(* IEC 61131-3 sources: plcassist-cli/packages/volt-lsp-iec/test-corpus/lenze-mid/Device/Plc Logic/Application/Library Manager/CommFB, 41 files *)

(* ---- ADDRESSCONCEPT.gvl ---- *)
VAR_GLOBAL
	DUMMY : UDINT := 0;
END_VAR

(* ---- CONSTANTS.gvl ---- *)
VAR_GLOBAL
	INVALID_ID : UDINT := 16#FFFFFFFF;
	MAX_PN_ALARM_DATA : UDINT := 198;
END_VAR

(* ---- ICOMMFBALARMSENDER.itf ---- *)
INTERFACE ICOMMFBALARMSENDER
END_INTERFACE

METHOD ALARMCNF
VAR_INPUT
	ERROR : DWORD;
END_VAR
END_METHOD

(* ---- ICOMMFBCONNECTIONMANAGERFACTORY.itf ---- *)
INTERFACE ICOMMFBCONNECTIONMANAGERFACTORY
END_INTERFACE

METHOD GETCONNECTIONMANAGER : UDINT
VAR_INPUT
	CLIENT : IConnectionManagerClient;
END_VAR
VAR_OUTPUT
	CONNECTIONMANAGER : IConnectionManager;
END_VAR
VAR_IN_OUT
	D_ADDR : ADDR_TYPE;
END_VAR
END_METHOD

METHOD RELEASECONNECTIONMANAGER : UDINT
VAR_INPUT
	CLIENT : IConnectionManagerClient;
	CONNECTIONMANAGER : IConnectionManager;
END_VAR
END_METHOD

(* ---- ICOMMFBDIAGPROVIDER.itf ---- *)
INTERFACE ICOMMFBDIAGPROVIDER
END_INTERFACE

METHOD CHECKOWNER : BOOL
VAR_INPUT
	ID : UDINT;
END_VAR
END_METHOD

METHOD GETALARM : DWORD
VAR_INPUT
	MODE : INT;
	F_ID : DWORD;
END_VAR
VAR_OUTPUT
	NEW : BOOL;
	ID : DWORD;
	LEN : INT;
END_VAR
VAR_IN_OUT
	AINFO : AINFO_TYPE;
	CURRENTALARMID : UDINT;
END_VAR
END_METHOD

METHOD GETDIAG : DWORD
VAR_INPUT
	ID : DWORD;
END_VAR
VAR_OUTPUT
	BUSY : BOOL;
	LEN : INT;
END_VAR
VAR_IN_OUT
	DINFO : DP_DIAG;
END_VAR
END_METHOD

(* ---- ICOMMFBFACTORY.itf ---- *)
INTERFACE ICOMMFBFACTORY
END_INTERFACE

METHOD CHECKOWNER : BOOL
VAR_INPUT
	ID : UDINT;
END_VAR
END_METHOD

METHOD GETRDREC : POINTER TO RDRECBase
VAR_INPUT
	ID : UDINT;
END_VAR
VAR_IN_OUT
	CLIENT : RDREC;
END_VAR
END_METHOD

METHOD GETWRREC : POINTER TO WRRECBase
VAR_INPUT
	ID : UDINT;
END_VAR
VAR_IN_OUT
	CLIENT : WRREC;
END_VAR
END_METHOD

METHOD RELEASERDREC : BOOL
VAR_INPUT
	ID : UDINT;
END_VAR
VAR_IN_OUT
	CLIENT : RDREC;
END_VAR
END_METHOD

METHOD RELEASEWRREC : BOOL
VAR_INPUT
	ID : UDINT;
END_VAR
VAR_IN_OUT
	CLIENT : WRREC;
END_VAR
END_METHOD

(* ---- ICOMMFBFACTORYEXT.itf ---- *)
INTERFACE ICOMMFBFACTORYEXT
END_INTERFACE

METHOD TRYGETADDRESS : BOOL
VAR_INPUT
	ID : DWORD;
END_VAR
VAR_OUTPUT
	STATUS : DWORD;
END_VAR
VAR_IN_OUT
	ADDR : ADDR_TYPE;
END_VAR
END_METHOD

METHOD TRYGETID : BOOL
VAR_OUTPUT
	STATUS : DWORD;
	ID : DWORD;
END_VAR
VAR_IN_OUT
	ADDR : ADDR_TYPE;
END_VAR
END_METHOD

(* ---- ICOMMFBFACTORYIO.itf ---- *)
INTERFACE ICOMMFBFACTORYIO
END_INTERFACE

METHOD CHECKOWNER : BOOL
VAR_INPUT
	ID : UDINT;
END_VAR
END_METHOD

METHOD GETINPUTDATA : DWORD
VAR_INPUT
	ID : DWORD;
	OFFSET : UINT;
	LEN : UINT;
	INPUTS : POINTER TO BYTE;
END_VAR
VAR_OUTPUT
	IO_LEN : UINT;
	CONSISTENCY : BOOL;
END_VAR
END_METHOD

METHOD PUTOUTPUTDATA : DWORD
VAR_INPUT
	ID : DWORD;
	OFFSET : UINT;
	LEN : UINT;
	OUTPUTS : POINTER TO BYTE;
END_VAR
VAR_OUTPUT
	IO_LEN : UINT;
	CONSISTENCY : BOOL;
END_VAR
END_METHOD

(* ---- ICOMMFBFIELDDEVICE.itf ---- *)
INTERFACE ICOMMFBFIELDDEVICE
END_INTERFACE

METHOD ALARMREQ : DWORD
VAR_INPUT
	ALARMSENDER : ICommFBAlarmSender;
	ID : DWORD;
	ATYPE : UINT;
	ASPEC : UINT;
	LEN : UINT;
	AINFO : POINTER TO BYTE;
END_VAR
END_METHOD

METHOD CHECKREADIND : BOOL
VAR_INPUT
	MODE : UINT;
	F_ID : DWORD;
END_VAR
VAR_OUTPUT
	STATUS : DWORD;
	IND : Read_Ind;
END_VAR
END_METHOD

METHOD CHECKWRITEIND : BOOL
VAR_INPUT
	MODE : UINT;
	F_ID : DWORD;
END_VAR
VAR_OUTPUT
	STATUS : DWORD;
	IND : Write_Ind;
END_VAR
END_METHOD

METHOD READNEGRSP : DWORD
VAR_INPUT
	CODE1 : BYTE;
	CODE2 : BYTE;
END_VAR
VAR_IN_OUT
	IND : Read_Ind;
END_VAR
END_METHOD

METHOD READRSP : DWORD
VAR_INPUT
	LEN : UINT;
	RECORD : POINTER TO BYTE;
END_VAR
VAR_IN_OUT
	IND : Read_Ind;
END_VAR
END_METHOD

METHOD WRITENEGRSP : DWORD
VAR_INPUT
	CODE1 : BYTE;
	CODE2 : BYTE;
END_VAR
VAR_IN_OUT
	IND : Write_Ind;
END_VAR
END_METHOD

METHOD WRITERSP : DWORD
VAR_IN_OUT
	IND : Write_Ind;
END_VAR
END_METHOD

(* ---- ICONNECTIONMANAGER.itf ---- *)
INTERFACE ICONNECTIONMANAGER
END_INTERFACE

METHOD CONNECTREQ : DWORD
VAR_IN_OUT
	D_ADDR : ADDR_TYPE;
END_VAR
END_METHOD

METHOD RELEASEREQ : DWORD
END_METHOD

METHOD UPDATEADDRESS : DWORD
VAR_IN_OUT
	D_ADDR : ADDR_TYPE;
END_VAR
END_METHOD

(* ---- ICONNECTIONMANAGERCLIENT.itf ---- *)
INTERFACE ICONNECTIONMANAGERCLIENT
END_INTERFACE

METHOD CONNECTCNF
VAR_INPUT
	ID : DWORD;
	ERRORCODE : DWORD;
END_VAR
END_METHOD

METHOD ERRORIND
VAR_INPUT
	ERRORCODE : DWORD;
END_VAR
END_METHOD

METHOD RELEASECNF
VAR_INPUT
	ERRORCODE : DWORD;
END_VAR
END_METHOD

(* ---- IGENERICIDFACTORY.itf ---- *)
INTERFACE IGENERICIDFACTORY
END_INTERFACE

METHOD TRYGETIDFROMREFERENCE : BOOL
VAR_INPUT
	PREF : POINTER TO BYTE;
END_VAR
VAR_OUTPUT
	ID : DWORD;
END_VAR
END_METHOD

(* ---- ADDR.fun ---- *)
FUNCTION ADDR : DWORD
VAR_INPUT
	EN : BOOL := TRUE;
	ID : DWORD;
END_VAR
VAR_OUTPUT
	ENO : BOOL;
END_VAR
END_FUNCTION

(* ---- GETLIBVERSION.fun ---- *)
FUNCTION GETLIBVERSION : VERSION
END_FUNCTION

(* ---- GETLIBVERSIONNUMBER.fun ---- *)
FUNCTION GETLIBVERSIONNUMBER : DWORD
END_FUNCTION

(* ---- ID.fun ---- *)
FUNCTION ID : DWORD
VAR_INPUT
	EN : BOOL := TRUE;
	MASTER : BYTE;
	SEGMENT : BYTE;
	STATION : BYTE;
	SLOT : BYTE;
END_VAR
END_FUNCTION

(* ---- ID_FROM_REF.fun ---- *)
FUNCTION ID_FROM_REF : DWORD
VAR_INPUT
	PREF : POINTER TO BYTE;
END_VAR
END_FUNCTION

(* ---- ISLIBRELEASED.fun ---- *)
FUNCTION ISLIBRELEASED : BOOL
END_FUNCTION

(* ---- SLOT_ID.fun ---- *)
FUNCTION SLOT_ID : DWORD
VAR_INPUT
	EN : BOOL := TRUE;
	ID : DWORD;
	SLOT : BYTE;
END_VAR
VAR_OUTPUT
	ENO : BOOL;
END_VAR
END_FUNCTION

(* ---- SUBSLOT_ID.fun ---- *)
FUNCTION SUBSLOT_ID : DWORD
VAR_INPUT
	EN : BOOL := TRUE;
	ID : DWORD;
	SLOT : UINT;
	SUBSLOT : UINT;
END_VAR
VAR_OUTPUT
	ENO : BOOL;
END_VAR
END_FUNCTION

(* ---- ADDR_TO_ID.fb ---- *)
FUNCTION_BLOCK ADDR_TO_ID
VAR_INPUT
	EN : BOOL := TRUE;
END_VAR
VAR_OUTPUT
	ENO : BOOL;
	STATUS : DWORD;
	ID : DWORD;
END_VAR
VAR_IN_OUT
	ADDR : ADDR_TYPE;
END_VAR
VAR
	S_INSTANCEHANDLER : InstanceHandler;
	I : DINT;
END_VAR
END_FUNCTION_BLOCK

(* ---- ALARMSENDERINTERNAL.fb ---- *)
FUNCTION_BLOCK ALARMSENDERINTERNAL
VAR_INPUT
	SALARM : POINTER TO SALARM;
END_VAR
END_FUNCTION_BLOCK

METHOD ALARMCNF
VAR_INPUT
	ERROR : DWORD;
END_VAR
END_METHOD

(* ---- CNCT.fb ---- *)
FUNCTION_BLOCK CNCT
VAR_INPUT
	REQ : BOOL;
	D_ADDR : ADDR_TYPE;
END_VAR
VAR_OUTPUT
	VALID : BOOL;
	ERROR : BOOL;
	BUSY : BOOL;
	STATUS : DWORD;
	ID : DWORD := Constants.INVALID_ID;
END_VAR
VAR
	S_INSTANCEHANDLER : InstanceHandler;
	_FACTORY : ICommFBConnectionManagerFactory;
	_CONNECTIONMANAGER : IConnectionManager;
	_REQ : BOOL;
	_STATE : CNCT_State := CNCT_State.S2_Idle;
	_ERRORCODE : UDINT;
	_CONNECTREQ : UDINT;
	_CONNECTID : DWORD := Constants.INVALID_ID;
	_RECVCONNECTCNF : BOOL;
	_RECVRELEASECNF : BOOL;
	_RECVABORTIND : BOOL;
	_CLIENT : ConnectionManagerClientInternal;
END_VAR
END_FUNCTION_BLOCK

METHOD ABORTIND
VAR_INPUT
	ERRORCODE : DWORD;
END_VAR
END_METHOD

METHOD CONNECTCNF
VAR_INPUT
	ID : DWORD;
	ERRORCODE : DWORD;
END_VAR
END_METHOD

METHOD RELEASECNF
VAR_INPUT
	ERRORCODE : DWORD;
END_VAR
END_METHOD

(* ---- CONNECTIONMANAGERCLIENTIMPLICITID.fb ---- *)
FUNCTION_BLOCK CONNECTIONMANAGERCLIENTIMPLICITID
VAR_INPUT
	CNCT : POINTER TO CREATE_ID;
END_VAR
END_FUNCTION_BLOCK

METHOD CONNECTCNF
VAR_INPUT
	ID : DWORD;
	ERRORCODE : DWORD;
END_VAR
END_METHOD

METHOD ERRORIND
VAR_INPUT
	ERRORCODE : DWORD;
END_VAR
END_METHOD

METHOD RELEASECNF
VAR_INPUT
	ERRORCODE : DWORD;
END_VAR
END_METHOD

(* ---- CONNECTIONMANAGERCLIENTINTERNAL.fb ---- *)
FUNCTION_BLOCK CONNECTIONMANAGERCLIENTINTERNAL
VAR_INPUT
	CNCT : POINTER TO CNCT;
END_VAR
END_FUNCTION_BLOCK

METHOD CONNECTCNF
VAR_INPUT
	ID : DWORD;
	ERRORCODE : DWORD;
END_VAR
END_METHOD

METHOD ERRORIND
VAR_INPUT
	ERRORCODE : DWORD;
END_VAR
END_METHOD

METHOD RELEASECNF
VAR_INPUT
	ERRORCODE : DWORD;
END_VAR
END_METHOD

(* ---- CREATE_ID.fb ---- *)
FUNCTION_BLOCK CREATE_ID
VAR_INPUT
	EN : BOOL := TRUE;
END_VAR
VAR_OUTPUT
	ENO : BOOL;
	STATUS : DWORD;
	ID : DWORD;
END_VAR
VAR_IN_OUT
	ADDR : ADDR_TYPE;
END_VAR
VAR
	S_INSTANCEHANDLER : InstanceHandler;
	_FACTORY : ICommFBConnectionManagerFactory;
	_CONNECTIONMANAGER : IConnectionManager;
	_STATE : CNCT_State := CNCT_State.S2_Idle;
	_ERRORCODE : UDINT;
	_CONNECTID : DWORD := Constants.INVALID_ID;
	_RECVCONNECTCNF : BOOL;
	_RECVRELEASECNF : BOOL;
	_RECVABORTIND : BOOL;
	_CLIENT : ConnectionManagerClientImplicitID;
	D_ADDR : ADDR_TYPE;
END_VAR
END_FUNCTION_BLOCK

METHOD ABORTIND
VAR_INPUT
	ERRORCODE : DWORD;
END_VAR
END_METHOD

METHOD CONNECTCNF
VAR_INPUT
	ID : DWORD;
	ERRORCODE : DWORD;
END_VAR
END_METHOD

METHOD RELEASECNF
VAR_INPUT
	ERRORCODE : DWORD;
END_VAR
END_METHOD

(* ---- GETIO_PART.fb ---- *)
FUNCTION_BLOCK GETIO_PART
VAR_INPUT
	EN : BOOL;
	ID : DWORD;
	OFFSET : INT;
	LEN : INT;
	INPUTS : POINTER TO BYTE;
END_VAR
VAR_OUTPUT
	ENO : BOOL;
	STATUS : DWORD;
	ERROR : BOOL;
END_VAR
VAR
	S_INSTANCEHANDLER : InstanceHandler;
	I : DINT;
	_FACTORY : ICommFBFactoryIO;
	IOLEN : UINT;
	TRANSFERCONSISTENT : BOOL;
END_VAR
END_FUNCTION_BLOCK

(* ---- ID_TO_ADDR.fb ---- *)
FUNCTION_BLOCK ID_TO_ADDR
VAR_INPUT
	EN : BOOL := TRUE;
	ID : DWORD;
END_VAR
VAR_OUTPUT
	ENO : BOOL;
	STATUS : DWORD;
END_VAR
VAR_IN_OUT
	ADDR : ADDR_TYPE;
END_VAR
VAR
	S_INSTANCEHANDLER : InstanceHandler;
	I : DINT;
	FACTORY : ICommFBFactoryExt;
END_VAR
END_FUNCTION_BLOCK

(* ---- INSTANCEHANDLER.fb ---- *)
FUNCTION_BLOCK INSTANCEHANDLER
VAR
	S_INSTANCECOUNT : UINT;
	S_FACTORIES : ARRAY [0..(MAX_INSTANCES - 1)] OF ICommFBFactory;
	S_FACTORIESEXT : ARRAY [0..(MAX_INSTANCES - 1)] OF ICommFBFactoryExt;
	S_FACTORIESIO : ARRAY [0..(MAX_INSTANCES - 1)] OF ICommFBFactoryIO;
	S_FACTORIESCONNECTIONS : ARRAY [0..(MAX_INSTANCES - 1)] OF ICommFBConnectionManagerFactory;
	S_FIELDDEVICES : ARRAY [0..(MAX_INSTANCES - 1)] OF ICommFBFieldDevice;
	S_GENERICIDFACTORIES : ARRAY [0..(MAX_INSTANCES - 1)] OF IGenericIDFactory;
	S_IDS : UDINT := (MAX_INSTANCES - 1);
	S_DIAGPROVIDERS : ARRAY [0..(MAX_INSTANCES - 1)] OF ICommFBDiagProvider;
	MAX_INSTANCES : UINT := 8;
END_VAR
END_FUNCTION_BLOCK

METHOD CREATEID : UDINT
END_METHOD

METHOD GETCONNECTIONMANAGERFACTORY : UDINT
VAR_OUTPUT
	FACTORY : ICommFBConnectionManagerFactory;
END_VAR
VAR_IN_OUT
	D_ADDR : ADDR_TYPE;
END_VAR
END_METHOD

METHOD GETDIAGFACTORY : UDINT
VAR_INPUT
	ID : UDINT;
END_VAR
VAR_OUTPUT
	DIAGPROVIDER : ICommFBDiagProvider;
END_VAR
END_METHOD

METHOD GETFACTORY : ICommFBFactory
VAR_INPUT
	ID : UDINT;
END_VAR
END_METHOD

METHOD GETFIELDDEVICE : DWORD
VAR_INPUT
	ID : UDINT;
END_VAR
VAR_OUTPUT
	FIELDDEVICE : ICommFBFieldDevice;
END_VAR
END_METHOD

METHOD GETIOFACTORY : UDINT
VAR_INPUT
	ID : UDINT;
END_VAR
VAR_OUTPUT
	FACTORY : ICommFBFactoryIO;
END_VAR
END_METHOD

METHOD REGISTER : UINT
VAR_INPUT
	FACTORY : ICommFBFactory;
END_VAR
END_METHOD

METHOD REGISTERDIAG : UINT
VAR_INPUT
	FACTORY : ICommFBFactory;
	DIAGPROVIDER : ICommFBDiagProvider;
END_VAR
END_METHOD

METHOD REGISTEREXT : UINT
VAR_INPUT
	FACTORY : ICommFBFactory;
	DIAGPROVIDER : ICommFBDiagProvider;
	FACTORYEXT : ICommFBFactoryExt;
END_VAR
END_METHOD

METHOD REGISTEREXTIO : UINT
VAR_INPUT
	FACTORY : ICommFBFactory;
	DIAGPROVIDER : ICommFBDiagProvider;
	FACTORYEXT : ICommFBFactoryExt;
	UPDATEIO : ICommFBFactoryIO;
END_VAR
END_METHOD

METHOD REGISTERFIELDDEVICE : UINT
VAR_INPUT
	FACTORY : ICommFBFactory;
	FACTORYEXT : ICommFBFactoryExt;
	DEVICE : ICommFBFieldDevice;
END_VAR
END_METHOD

METHOD REGISTERINTERFACES : UINT
VAR_INPUT
	FACTORY : ICommFBFactory;
	DIAGPROVIDER : ICommFBDiagProvider;
	FACTORYEXT : ICommFBFactoryExt;
	UPDATEIO : ICommFBFactoryIO;
	CNCT : ICommFBConnectionManagerFactory;
END_VAR
END_METHOD

(* ---- PRVREC.fb ---- *)
FUNCTION_BLOCK PRVREC
VAR_INPUT
	EN : BOOL;
	MODE : UINT;
	F_ID : DWORD;
	CODE1 : BYTE;
	CODE2 : BYTE;
	LEN : UINT;
	RECORD : POINTER TO BYTE;
END_VAR
VAR_OUTPUT
	ENO : BOOL;
	NEW : BOOL;
	STATUS : DWORD;
	SLOT : UINT;
	SUBSLOT : UINT;
	INDEX : UINT;
	RLEN : UINT;
END_VAR
VAR
	S_INSTANCEHANDLER : InstanceHandler;
	_STATE : PRVREC_State := PRVREC_State.S1_INIT;
	_DEVICE : ICommFBFieldDevice;
	_READIND : Read_Ind;
	EMPTYIND : Read_Ind;
END_VAR
END_FUNCTION_BLOCK

(* ---- RALARM.fb ---- *)
FUNCTION_BLOCK RALARM
VAR_INPUT
	EN : BOOL;
	MODE : INT;
	F_ID : DWORD;
END_VAR
VAR_OUTPUT
	ENO : BOOL;
	NEW : BOOL;
	STATUS : DWORD;
	ID : DWORD;
	LEN : INT;
END_VAR
VAR_IN_OUT
	AINFO : AINFO_TYPE;
END_VAR
VAR
	S_INSTANCEHANDLER : InstanceHandler;
	M_EN : BOOL;
	M_MODE : INT;
	M_F_ID : DWORD;
	M_FACTORY : ICommFBDiagProvider;
	M_CURRENTALARMID : UDINT := Constants.INVALID_ID;
END_VAR
END_FUNCTION_BLOCK

(* ---- RCVREC.fb ---- *)
FUNCTION_BLOCK RCVREC
VAR_INPUT
	EN : BOOL;
	MODE : UINT;
	F_ID : DWORD;
	MLEN : UINT;
	CODE1 : BYTE;
	CODE2 : BYTE;
	RECORD : POINTER TO BYTE;
END_VAR
VAR_OUTPUT
	ENO : BOOL;
	NEW : BOOL;
	STATUS : DWORD;
	SLOT : UINT;
	SUBSLOT : UINT;
	INDEX : UINT;
	LEN : UINT;
END_VAR
VAR
	S_INSTANCEHANDLER : InstanceHandler;
	_STATE : RCVREC_State := RCVREC_State.S1_INIT;
	_DEVICE : ICommFBFieldDevice;
	_WRITEIND : Write_Ind;
	EMPTYIND : Write_Ind;
	I : DINT;
END_VAR
END_FUNCTION_BLOCK

(* ---- RDIAG.fb ---- *)
FUNCTION_BLOCK RDIAG
VAR_INPUT
	REQ : BOOL;
	ID : DWORD;
	MLEN : INT;
END_VAR
VAR_OUTPUT
	VALID : BOOL;
	BUSY : BOOL;
	ERROR : BOOL;
	STATUS : DWORD;
	LEN : INT;
END_VAR
VAR_IN_OUT
	DINFO : DP_DIAG;
END_VAR
VAR
	S_INSTANCEHANDLER : InstanceHandler;
	M_FACTORY : ICommFBDiagProvider;
END_VAR
END_FUNCTION_BLOCK

(* ---- RDREC.fb ---- *)
FUNCTION_BLOCK RDREC
VAR_INPUT
	REQ : BOOL;
	ID : DWORD;
	INDEX : INT;
	MLEN : INT;
	RECORD : POINTER TO BYTE;
END_VAR
VAR_OUTPUT
	VALID : BOOL;
	BUSY : BOOL;
	ERROR : BOOL;
	STATUS : DWORD;
	LEN : INT;
END_VAR
VAR
	M_FACTORY : ICommFBFactory;
	M_PRDREC : POINTER TO RDRECbase;
	_REQ : BOOL;
	S_INSTANCEHANDLER : InstanceHandler;
END_VAR
END_FUNCTION_BLOCK

(* ---- RDRECBASE.fb ---- *)
FUNCTION_BLOCK RDRECBASE
VAR_INPUT
	REQ : BOOL;
	ID : DWORD;
	INDEX : INT;
	MLEN : INT;
	RECORD : POINTER TO BYTE;
END_VAR
VAR_OUTPUT
	VALID : BOOL;
	ERROR : BOOL;
	BUSY : BOOL;
	STATUS : DWORD;
	LEN : INT;
END_VAR
END_FUNCTION_BLOCK

(* ---- RDRECDEFAULT.fb ---- *)
FUNCTION_BLOCK RDRECDEFAULT EXTENDS RDRECbase
VAR
	STATE : RDREC_State := RDREC_State.S2_Idle;
	_ERRORCODE : UDINT;
	DATALEN : INT;
	PRECORDDATA : POINTER TO BYTE;
	NEXT : BOOL;
END_VAR
END_FUNCTION_BLOCK

METHOD COPYDATA
VAR_INPUT
	LENGTH : INT;
	PDATA : POINTER TO BYTE;
END_VAR
END_METHOD

METHOD NEGRESPONSE
VAR_INPUT
	ERRORCODE : DWORD;
END_VAR
END_METHOD

METHOD POSRESPONSE
END_METHOD

METHOD START : UDINT
END_METHOD

METHOD WAITING
END_METHOD

(* ---- SALARM.fb ---- *)
FUNCTION_BLOCK SALARM
VAR_INPUT
	REQ : BOOL;
	ID : DWORD;
	ATYPE : UINT;
	ASPEC : UINT;
	LEN : UINT;
	AINFO : POINTER TO BYTE;
END_VAR
VAR_OUTPUT
	DONE : BOOL;
	BUSY : BOOL;
	ERROR : BOOL;
	STATUS : DWORD;
END_VAR
VAR
	S_INSTANCEHANDLER : InstanceHandler;
	_REQ : BOOL;
	_STATE : SALRM_State := SALRM_State.S1_INIT;
	SEND_RESULT : UDINT;
	_DEVICE : ICommFBFieldDevice;
	_CLIENT : AlarmSenderInternal;
	_ERROR : DWORD;
	_CONTINUE : BOOL;
END_VAR
END_FUNCTION_BLOCK

METHOD ALARMCNF
VAR_INPUT
	ERROR : DWORD;
END_VAR
END_METHOD

METHOD NEG_RESPONSE
VAR_INPUT
	ERROR : DWORD;
END_VAR
END_METHOD

METHOD POS_RESPONSE
END_METHOD

(* ---- SETIO_PART.fb ---- *)
FUNCTION_BLOCK SETIO_PART
VAR_INPUT
	EN : BOOL;
	ID : DWORD;
	OFFSET : INT;
	LEN : INT;
	OUTPUTS : POINTER TO BYTE;
END_VAR
VAR_OUTPUT
	ENO : BOOL;
	STATUS : DWORD;
	ERROR : BOOL;
END_VAR
VAR
	S_INSTANCEHANDLER : InstanceHandler;
	I : DINT;
	_FACTORY : ICommFBFactoryIO;
	IOLEN : UINT;
	TRANSFERCONSISTENT : BOOL;
END_VAR
END_FUNCTION_BLOCK

(* ---- WRREC.fb ---- *)
FUNCTION_BLOCK WRREC
VAR_INPUT
	REQ : BOOL;
	ID : DWORD;
	INDEX : INT;
	LEN : INT;
	RECORD : POINTER TO BYTE;
END_VAR
VAR_OUTPUT
	DONE : BOOL;
	BUSY : BOOL;
	ERROR : BOOL;
	STATUS : DWORD;
END_VAR
VAR
	M_FACTORY : ICommFBFactory;
	M_PWRREC : POINTER TO WRRECbase;
	_REQ : BOOL;
	S_INSTANCEHANDLER : InstanceHandler;
END_VAR
END_FUNCTION_BLOCK

(* ---- WRRECBASE.fb ---- *)
FUNCTION_BLOCK WRRECBASE
VAR_INPUT
	REQ : BOOL;
	ID : DWORD;
	INDEX : INT;
	LEN : INT;
	RECORD : POINTER TO BYTE;
END_VAR
VAR_OUTPUT
	DONE : BOOL;
	BUSY : BOOL;
	ERROR : BOOL;
	STATUS : DWORD;
END_VAR
END_FUNCTION_BLOCK

(* ---- WRRECDEFAULT.fb ---- *)
FUNCTION_BLOCK WRRECDEFAULT EXTENDS WRRECbase
VAR
	STATE : WRREC_State := WRREC_State.S2_Idle;
	ERRORCODE : UDINT;
END_VAR
END_FUNCTION_BLOCK

METHOD NEGRESPONSE
VAR_INPUT
	ERRORCODE : DWORD;
END_VAR
END_METHOD

METHOD POSRESPONSE
END_METHOD

METHOD START : UDINT
END_METHOD

METHOD WAITING
END_METHOD
